(* IEC 61131-3 sources: plc-st-coding-agent/progress/f14_agent_v2/release/datasets/public/tests, 20 files *)

(* ---- public-easy-01.reference.st ---- *)
(* 参考解：Automated filling line control（清洗 -> 灌装 -> 压盖 -> 包装 -> 完成灯 -> 取瓶复位）
   工序号用内部状态 stepNo 表示：0=空闲 1=清洗 2=灌装 3=压盖 4=包装 5=完成。
   只用接口变量做输出，“工序启动后保持运行”由 stepNo 只增不减保证。 *)
FUNCTION_BLOCK FB_FillingLine
VAR_INPUT
    bottleSensor : BOOL;            (* 瓶子到位检测 *)
    cleaningConfirmButton : BOOL;   (* 清洗完成确认 *)
    fillingConfirmButton : BOOL;    (* 灌装完成确认 *)
    cappingConfirmButton : BOOL;    (* 压盖完成确认 *)
    packingConfirmButton : BOOL;    (* 包装完成确认 *)
    finishedButton : BOOL;          (* 取走瓶子确认 *)
END_VAR
VAR_OUTPUT
    Pump_Motor : BOOL;              (* 清洗泵 *)
    Filling_Valve : BOOL;           (* 灌装阀 *)
    Capping_Machine : BOOL;         (* 压盖机 *)
    Packing_Machine : BOOL;         (* 包装机 *)
    Completion_Light : BOOL;        (* 包装完成指示灯 *)
END_VAR
VAR
    stepNo : INT;                   (* 当前工序号，0=空闲 *)
END_VAR

(* R1: 检测到瓶子就启动清洗泵（stepNo 1），此后 stepNo 不回退，泵持续工作 *)
IF bottleSensor AND (stepNo = 0) THEN
    stepNo := 1;
END_IF

(* R2..R5: 每道工序由“上一道工序完成”的确认按钮推进；只接受当拍工序的确认，
   因此误按后道工序的按钮不会跳步，而且机器一旦启动就保持运行 *)
IF (stepNo = 1) AND cleaningConfirmButton THEN
    stepNo := 2;
ELSIF (stepNo = 2) AND fillingConfirmButton THEN
    stepNo := 3;
ELSIF (stepNo = 3) AND cappingConfirmButton THEN
    stepNo := 4;
ELSIF (stepNo = 4) AND packingConfirmButton THEN
    stepNo := 5;
END_IF

(* R6: 取走瓶子 -> 灭灯并整线复位，准备下一循环 *)
IF finishedButton THEN
    stepNo := 0;
END_IF

(* 各执行机构的输出：由工序号唯一决定，故“启动即保持” *)
Pump_Motor := (stepNo >= 1);
Filling_Valve := (stepNo >= 2);
Capping_Machine := (stepNo >= 3);
Packing_Machine := (stepNo >= 4);
Completion_Light := (stepNo = 5);
END_FUNCTION_BLOCK

(* ---- public-easy-02.reference.st ---- *)
(* 参考解：Dual-word edge detection（DWORD 逐位上升沿/下降沿）
   prevValue 保存上一拍的输入值，声明初值为 0（PLC 上电瞬间存储区为 0），
   因此第 1 拍等价于“相对全 0 的边沿检测”，与需求“比较两个连续的 DWORD”一致。 *)
FUNCTION_BLOCK FB_DualWordEdge
VAR_INPUT
    value : DWORD;                  (* 每个周期检查的输入字 *)
END_VAR
VAR_OUTPUT
    hasChanged : BOOL;              (* 有无任何位变化 *)
    hasRisingEdges : BOOL;          (* 有无上升沿 *)
    risingBits : DWORD;             (* 上升沿位流：某位本拍由 0 变 1 则为 1 *)
    noOfRisingBits : USINT;         (* 上升沿位数 *)
    hasFallingEdges : BOOL;         (* 有无下降沿 *)
    fallingBits : DWORD;            (* 下降沿位流：某位本拍由 1 变 0 则为 1 *)
    noOfFallingBits : USINT;        (* 下降沿位数 *)
END_VAR
VAR
    prevValue : DWORD;              (* 上一拍的输入值 *)
    tmpBits : DWORD;                (* 统计位数的移位暂存 *)
    bitCount : USINT;               (* 统计结果暂存 *)
    i : INT;                        (* 循环变量 *)
END_VAR

(* R1/R2: 按位求差。NOT 对整数是 32 位按位取反，与 DWORD 宽度一致。
   IEC 的 AND/OR 两侧都是整数时按位运算，所以这里不会退化成逻辑运算。 *)
risingBits := value AND NOT prevValue;
fallingBits := prevValue AND NOT value;

(* R3: 是否变化，以及两类边沿是否存在 *)
hasChanged := (risingBits <> 0) OR (fallingBits <> 0);
hasRisingEdges := risingBits <> 0;
hasFallingEdges := fallingBits <> 0;

(* R4: 上升沿位数——逐位右移数 1 的个数（32 位，故循环 32 次） *)
bitCount := 0;
tmpBits := risingBits;
FOR i := 1 TO 32 DO
    IF (tmpBits AND 1) <> 0 THEN
        bitCount := bitCount + 1;
    END_IF
    tmpBits := tmpBits SHR 1;
END_FOR
noOfRisingBits := bitCount;

(* R6: 下降沿位数，同一套逐位统计 *)
bitCount := 0;
tmpBits := fallingBits;
FOR i := 1 TO 32 DO
    IF (tmpBits AND 1) <> 0 THEN
        bitCount := bitCount + 1;
    END_IF
    tmpBits := tmpBits SHR 1;
END_FOR
noOfFallingBits := bitCount;

(* R5: 本拍值成为下一拍的“上一拍” *)
prevValue := value;
END_FUNCTION_BLOCK

(* ---- public-easy-03.reference.st ---- *)
(* 参考解：Alarm handling（带回差的高/低限报警 + 参数校验）
   报警输出是锁存量：超过限值才置位，回到“限值 ± 回差”以内才复位（回差防抖）。
   参数非法时置 error 并给出 status，且本次扫描不再评估报警（等价于“退出程序”）。 *)
FUNCTION_BLOCK FB_AlarmHandling
VAR_INPUT
    Value : REAL;                   (* 被监视的输入值 *)
    hiLevel : REAL;                 (* 高限报警值 *)
    loLevel : REAL;                 (* 低限报警值 *)
    hystWindow : REAL;              (* 回差窗口 *)
END_VAR
VAR_OUTPUT
    hiAlarm : BOOL;                 (* 高限报警 *)
    loAlarm : BOOL;                 (* 低限报警 *)
    error : BOOL;                   (* 执行出错 *)
    status : WORD;                  (* 状态码：16#8001 / 16#8002 *)
END_VAR

(* R5: 上下限设置反了（loLevel >= hiLevel）-> error，status=16#8001，退出 *)
IF loLevel >= hiLevel THEN
    error := TRUE;
    status := 16#8001;
(* R6: 回差窗口不比正常范围窄（hystWindow >= hiLevel - loLevel）-> error，status=16#8002 *)
ELSIF hystWindow >= (hiLevel - loLevel) THEN
    error := TRUE;
    status := 16#8002;
ELSE
    error := FALSE;
    status := 16#0000;

    (* R1/R2: 高于高限置位；低于 hiLevel-hystWindow 才复位，中间的过渡带保持原状态 *)
    IF Value > hiLevel THEN
        hiAlarm := TRUE;
    ELSIF Value < (hiLevel - hystWindow) THEN
        hiAlarm := FALSE;
    END_IF

    (* R3/R4: 低于低限置位；高于 loLevel+hystWindow 才复位 *)
    IF Value < loLevel THEN
        loAlarm := TRUE;
    ELSIF Value > (loLevel + hystWindow) THEN
        loAlarm := FALSE;
    END_IF
END_IF
END_FUNCTION_BLOCK

(* ---- public-easy-04.reference.st ---- *)
FUNCTION_BLOCK FB
VAR_INPUT
    VISCOSITY_OK : BOOL;
    PASTE_E_STOP_NC : BOOL;
    DebounceTime : TIME;
    CycleTime : TIME;
END_VAR
VAR_OUTPUT
    VFD_RUN : BOOL;
    PUMP_MAINT_DUE : BOOL;
    PUMP_RUNTIME_ACC : LTIME;
END_VAR
VAR
    viscosityDelay : TON;
END_VAR
viscosityDelay(IN := VISCOSITY_OK AND PASTE_E_STOP_NC, PT := DebounceTime);
VFD_RUN := viscosityDelay.Q;
IF VFD_RUN THEN
    PUMP_RUNTIME_ACC := PUMP_RUNTIME_ACC + TIME_TO_LTIME(CycleTime);
END_IF;
PUMP_MAINT_DUE := PUMP_RUNTIME_ACC >= LTIME#500h;
END_FUNCTION_BLOCK

(* ---- public-easy-05.reference.st ---- *)
FUNCTION_BLOCK FB_WeldGapAlarm
VAR_INPUT
    Gap_Exceeded : BOOL;
    Weld_E_Stop_NC : BOOL;
    DebounceTime : TIME;
END_VAR
VAR_OUTPUT
    Operator_Alert : BOOL;
    Weld_Soft_Start_Active : BOOL;
END_VAR
VAR
    startupDelay : TON;
    gapDelay : TON;
END_VAR
startupDelay(IN := TRUE, PT := T#5s);
Weld_Soft_Start_Active := NOT startupDelay.Q;
gapDelay(IN := startupDelay.Q AND Weld_E_Stop_NC AND Gap_Exceeded, PT := DebounceTime);
Operator_Alert := gapDelay.Q;
END_FUNCTION_BLOCK

(* ---- public-easy-06.reference.st ---- *)
FUNCTION_BLOCK FB_AerationBlower
VAR_INPUT
    DO_LOW : BOOL;
    AERATION_E_STOP_NC : BOOL;
END_VAR
VAR_OUTPUT
    BLOWER_RUN : BOOL;
    AERATION_BLOWER_CYCLE_COUNT : UINT;
END_VAR
VAR
    startDelay : TON;
    wasRunning : BOOL;
END_VAR
startDelay(IN := DO_LOW AND AERATION_E_STOP_NC, PT := T#5s);
BLOWER_RUN := startDelay.Q;
IF BLOWER_RUN AND NOT wasRunning AND AERATION_BLOWER_CYCLE_COUNT < 65535 THEN
    AERATION_BLOWER_CYCLE_COUNT := AERATION_BLOWER_CYCLE_COUNT + 1;
END_IF;
wasRunning := BLOWER_RUN;
END_FUNCTION_BLOCK

(* ---- public-hard-01.reference.st ---- *)
(*
    public-hard-01  Material Proportioning Process Control
    参考解：单个 FUNCTION_BLOCK。接口名与数据类型严格照抄 variables。

    平台说明（公共题制作约定 §7）：
      * 无 TON / R_TRIG，按钮的上升沿用显式边沿
            e := btn AND NOT prev;  prev := btn;
        在扫描末尾统一滚动 prev，避免同拍重复触发。
      * "液位达到 N cm" 用 levelSensor >= N 判断（液位单调上升的语义）。
      * 时间类原语里没有可用的定时器，本题流程全部由 levelSensor / 完成信号推进。

    本文件用 (* R1: ... *) 形式标注需求编号，逐条对应 requirements。
*)
FUNCTION_BLOCK FB_MaterialProportioning
VAR_INPUT
    estop : BOOL;             (* R1 急停：FALSE = 触发 *)
    opeMode : BOOL;           (* R2/R4 运行方式：FALSE = 手动，TRUE = 自动 *)
    valveAStart : BOOL;       (* 手动按钮（上升沿启停） *)
    valveBStart : BOOL;
    valveCStart : BOOL;
    valveDStart : BOOL;
    mixMotorStart : BOOL;
    autoStart : BOOL;         (* 自动流程启动按钮（上升沿） *)
    processMode : BOOL;       (* R5 FALSE = 直接混合；TRUE = 先进 C 到 100cm 再混合 *)
    levelSensor : INT;        (* 液位传感器，单位 cm *)
    mixMotorComplete : BOOL;  (* R6 混合完成信号 *)
END_VAR
VAR_OUTPUT
    valveARun : BOOL;
    valveBRun : BOOL;
    valveCRun : BOOL;
    valveDRun : BOOL;
    mixMotorRun : BOOL;
END_VAR
VAR
    (* 自动流程步序：0 空闲 / 10 进料 A / 20 进料 B / 35 进料 C / 40 混合 / 50 完成 *)
    state : INT;
    (* 各按钮与运行方式上一拍的值（显式边沿用） *)
    prevAutoStart : BOOL;
    prevValveAStart : BOOL;
    prevValveBStart : BOOL;
    prevValveCStart : BOOL;
    prevValveDStart : BOOL;
    prevMixMotorStart : BOOL;
    prevOpeMode : BOOL;
    (* 手动模式下五个设备的启停记忆 *)
    manA : BOOL;
    manB : BOOL;
    manC : BOOL;
    manD : BOOL;
    manMix : BOOL;
END_VAR

(* R1: 急停最高优先级——estop=FALSE 时所有设备立即停机，
   并复位自动流程与手动记忆；急停解除后不会自动续跑，必须重新启动。 *)
IF NOT estop THEN
    state := 0;
    manA := FALSE;
    manB := FALSE;
    manC := FALSE;
    manD := FALSE;
    manMix := FALSE;
    valveARun := FALSE;
    valveBRun := FALSE;
    valveCRun := FALSE;
    valveDRun := FALSE;
    mixMotorRun := FALSE;

(* R2: 手动模式——五个设备各自由对应按钮的上升沿翻转（启/停）。
   R3: 只认上升沿：按住不放不会反复翻转；释放后保持当前状态。 *)
ELSIF NOT opeMode THEN
    (* 从自动切到手动的那一拍：放弃自动流程，手动记忆全部复位（需求未规定，
       取最安全侧，见文件末尾"需求未覆盖处"说明）。 *)
    IF prevOpeMode THEN
        state := 0;
        manA := FALSE;
        manB := FALSE;
        manC := FALSE;
        manD := FALSE;
        manMix := FALSE;
    END_IF
    IF valveAStart AND NOT prevValveAStart THEN
        manA := NOT manA;
    END_IF
    IF valveBStart AND NOT prevValveBStart THEN
        manB := NOT manB;
    END_IF
    IF valveCStart AND NOT prevValveCStart THEN
        manC := NOT manC;
    END_IF
    IF valveDStart AND NOT prevValveDStart THEN
        manD := NOT manD;
    END_IF
    IF mixMotorStart AND NOT prevMixMotorStart THEN
        manMix := NOT manMix;
    END_IF
    valveARun := manA;
    valveBRun := manB;
    valveCRun := manC;
    valveDRun := manD;
    mixMotorRun := manMix;

(* R4/R5/R6: 自动模式——按工艺步序推进设备，手动按钮被忽略。 *)
ELSE
    (* 刚进入自动模式：自动流程从头开始，手动残留输出全部关断。 *)
    IF NOT prevOpeMode THEN
        state := 0;
        valveARun := FALSE;
        valveBRun := FALSE;
        valveCRun := FALSE;
        valveDRun := FALSE;
        mixMotorRun := FALSE;
    END_IF

    CASE state OF
        0:  (* 空闲：等待 autoStart 上升沿 *)
            valveARun := FALSE;
            valveBRun := FALSE;
            valveCRun := FALSE;
            valveDRun := FALSE;
            mixMotorRun := FALSE;
            (* R4: 按 autoStart 启动自动流程，先开阀 A *)
            IF autoStart AND NOT prevAutoStart THEN
                state := 10;
                valveARun := TRUE;
            END_IF

        10: (* 进料 A：液位到 50cm 关 A、开 B *)
            valveARun := TRUE;
            valveBRun := FALSE;
            valveCRun := FALSE;
            valveDRun := FALSE;
            mixMotorRun := FALSE;
            IF levelSensor >= 50 THEN
                valveARun := FALSE;
                valveBRun := TRUE;
                state := 20;
            END_IF

        20: (* 进料 B：液位到 80cm 关 B；随后按 processMode 决定下一步 *)
            valveARun := FALSE;
            valveBRun := TRUE;
            valveCRun := FALSE;
            valveDRun := FALSE;
            mixMotorRun := FALSE;
            IF levelSensor >= 80 THEN
                valveBRun := FALSE;
                IF processMode THEN
                    (* R5(true): 先开 C 继续进料到 100cm *)
                    valveCRun := TRUE;
                    state := 35;
                ELSE
                    (* R5(false): 不进 C，直接启动混合电机 *)
                    mixMotorRun := TRUE;
                    state := 40;
                END_IF
            END_IF

        35: (* 进料 C：液位到 100cm 关 C、启动混合电机 *)
            valveARun := FALSE;
            valveBRun := FALSE;
            valveCRun := TRUE;
            valveDRun := FALSE;
            mixMotorRun := FALSE;
            IF levelSensor >= 100 THEN
                valveCRun := FALSE;
                mixMotorRun := TRUE;
                state := 40;
            END_IF

        40: (* 混合中：收到混合完成信号 → 停电机、开 D、流程结束 *)
            valveARun := FALSE;
            valveBRun := FALSE;
            valveCRun := FALSE;
            valveDRun := FALSE;
            mixMotorRun := TRUE;
            IF mixMotorComplete THEN
                mixMotorRun := FALSE;
                valveDRun := TRUE;
                state := 50;
            END_IF

        50: (* 完成：D 保持开启把料送出；再次 autoStart 开始新一周期 *)
            valveARun := FALSE;
            valveBRun := FALSE;
            valveCRun := FALSE;
            valveDRun := TRUE;
            mixMotorRun := FALSE;
            IF autoStart AND NOT prevAutoStart THEN
                valveDRun := FALSE;
                valveARun := TRUE;
                state := 10;
            END_IF
    END_CASE
END_IF

(* 边沿记忆统一在扫描末尾滚动（顺序不可提前，见约定 §7）。 *)
prevAutoStart := autoStart;
prevValveAStart := valveAStart;
prevValveBStart := valveBStart;
prevValveCStart := valveCStart;
prevValveDStart := valveDStart;
prevMixMotorStart := mixMotorStart;
prevOpeMode := opeMode;

(*
  需求未覆盖处的取舍（均为最安全侧，且已由 test_cases 覆盖其行为）：
  1) 运行方式切换：自动→手动或手动→自动时，当前流程被中止、输出全部关断，
     不会在切换后残留上一模式的设备动作；自动模式要从步序 0 重新 autoStart。
  2) 自动流程进行中再次按 autoStart 被忽略（按键只对步序 0 / 50 有效），
     避免运行中反复重启流程。
  3) 自动完成后阀 D 保持开启（"open valve D, and the automatic process ends"），
     直到下一次 autoStart 开始新周期或急停触发。
  4) 步序 0 与各步都显式给全部输出赋值，保证同一扫描周期内输出不残留上一步的值。
*)
END_FUNCTION_BLOCK

(* ---- public-hard-02.reference.st ---- *)
(* public-hard-02 Flexible Processing Control
   1# 上料 / 2#~4# 加工 / 5# 出库。工序序列由 processSequence + processLength 给出，
   processLength 从 processSequence[1] 起算，末项由 caller 保证是 5# 出库站。
   内部状态机 phase：0=空闲/待料，1=输送中，2=等当前加工工位完成信号。 *)

FUNCTION_BLOCK FB
VAR_INPUT
    processLength : USINT;
    sensor1 : BOOL;
    sensor2 : BOOL;
    sensor3 : BOOL;
    sensor4 : BOOL;
    sensor5 : BOOL;
    station1Start : BOOL;
    station2Complete : BOOL;
    station3Complete : BOOL;
    station4Complete : BOOL;
    processSequence : ARRAY[1..8] OF USINT;
END_VAR
VAR_OUTPUT
    conveyorLeft : BOOL;
    conveyorRight : BOOL;
END_VAR
VAR
    phase : INT;          (* 0 空闲；1 输送中；2 等加工完成 *)
    idx : INT;            (* 当前执行到 processSequence 的第几项 *)
    curStation : INT;     (* 产品当前所在工位 *)
    dstStation : INT;     (* 本段输送的目标工位 *)
    lenNow : INT;
    dstOK : BOOL;
    arrived : BOOL;
    startEdge : BOOL;
    startPrev : BOOL;
    compEdge : BOOL;
    comp2Prev : BOOL;
    comp3Prev : BOOL;
    comp4Prev : BOOL;
END_VAR

(* R1/R2: 启动按钮上升沿 + 1# 有料才启动；序列长度必须落在 1..8 *)
startEdge := station1Start AND NOT startPrev;
startPrev := station1Start;
lenNow := processLength;

(* 加工完成信号按上升沿消费；每拍都刷新历史值，避免边沿被相位切换吃掉 *)
compEdge := FALSE;
IF phase = 2 THEN
    IF curStation = 2 THEN
        compEdge := station2Complete AND NOT comp2Prev;
    ELSIF curStation = 3 THEN
        compEdge := station3Complete AND NOT comp3Prev;
    ELSIF curStation = 4 THEN
        compEdge := station4Complete AND NOT comp4Prev;
    END_IF;
END_IF;
comp2Prev := station2Complete;
comp3Prev := station3Complete;
comp4Prev := station4Complete;

conveyorLeft := FALSE;
conveyorRight := FALSE;

(* R1: 上料工位有料 + 按下启动 → 查第一个工序号，当拍就启动输送带 *)
IF phase = 0 THEN
    IF sensor1 AND startEdge THEN
        IF (lenNow >= 1) AND (lenNow <= 8) THEN
            dstStation := processSequence[1];
            dstOK := (dstStation >= 2) AND (dstStation <= 5);
            IF dstOK THEN
                idx := 1;
                curStation := 1;
                phase := 1;
            END_IF;
        END_IF;
    END_IF;
END_IF;

(* R4: 收到当前工位完成信号 → 查下一个工序号，当拍转向继续输送 *)
IF phase = 2 THEN
    IF compEdge THEN
        idx := idx + 1;
        IF (idx > lenNow) OR (idx > 8) THEN
            (* 非法序列（末项不是 5#）的保护：不再读数组下标，直接停机 *)
            phase := 0;
        ELSE
            dstStation := processSequence[idx];
            dstOK := (dstStation >= 2) AND (dstStation <= 5);
            IF dstOK THEN
                phase := 1;
            ELSE
                phase := 0;
            END_IF;
        END_IF;
    END_IF;
END_IF;

(* R3/R5: 按 "目标工位 vs 当前工位" 决定方向；只看目标工位传感器判到位 *)
IF phase = 1 THEN
    IF dstStation > curStation THEN
        conveyorRight := TRUE;
    ELSIF dstStation < curStation THEN
        conveyorLeft := TRUE;
    END_IF;
    arrived := FALSE;
    IF dstStation = 2 THEN
        arrived := sensor2;
    ELSIF dstStation = 3 THEN
        arrived := sensor3;
    ELSIF dstStation = 4 THEN
        arrived := sensor4;
    ELSIF dstStation = 5 THEN
        arrived := sensor5;
    END_IF;
    IF arrived THEN
        conveyorLeft := FALSE;
        conveyorRight := FALSE;
        curStation := dstStation;
        IF dstStation = 5 THEN
            (* R5: 送到 5# 出库站，一个产品的流程结束 *)
            phase := 0;
        ELSE
            (* R4: 停在该工位，等它给出加工完成信号 *)
            phase := 2;
        END_IF;
    END_IF;
END_IF;
END_FUNCTION_BLOCK

(* ---- public-hard-03.reference.st ---- *)
(*
  Recipe Management System — 参考解（public-hard-03）

  配方库 recipe 是 VAR_IN_OUT 的结构体数组，最多 10 条，recipeID = 0 表示空槽；
  四个请求信号取上升沿，因此一个请求只执行一次（电平保持不会重复执行）。

  需求编号（对应 requirements 的 Notes）：
    R2  查询：号码不存在 -> error=TRUE & status=16#8001；存在 -> 输出到 recipeQueryResult
    R3  新增：号码重复 -> 16#8002；无空槽 -> 16#8003；否则存到下标最小的空槽
    R4  删除：号码不存在 -> 16#8004；存在 -> 把该槽的 recipeID 置 0
    R5  修改：号码不存在 -> 16#8005；存在 -> 用 recipeIn 覆盖该槽
  另有 R1：配方字段 recipeID/ingredientType/ingredientRatio/productionTemperature。

  两处按需求原文做的判定口径（都写在下面的注释里）：
    * 0 号不是合法配方号：查询/删除/修改 0 号一律按"号码不存在"处理；
    * 新增时号码与本库任何一条 recipeID 相同即算重复，因此 0 号会与空槽的 0 相撞，
      在还有空槽时报 16#8002（R3 的判定顺序本来就是"先查重复、再查空槽"）。
*)

TYPE ST_Recipe :
STRUCT
  recipeID : INT;                (* 配方号，0 = 空槽 *)
  ingredientType : INT;          (* 原料类型 *)
  ingredientRatio : REAL;        (* 原料配比 *)
  productionTemperature : REAL;  (* 生产温度 *)
END_STRUCT
END_TYPE

FUNCTION_BLOCK FB
VAR_INPUT
  addRecipe : BOOL;              (* R3 新增请求 *)
  deleteRecipe : BOOL;           (* R4 删除请求 *)
  modifyRecipe : BOOL;           (* R5 修改请求 *)
  queryRecipe : BOOL;            (* R2 查询请求 *)
  recipeIn : ST_Recipe;          (* 请求携带的配方 *)
END_VAR
VAR_OUTPUT
  recipeAdded : BOOL;            (* 新增成功指示，只在执行成功那一拍为 TRUE *)
  recipeDeleted : BOOL;          (* 删除成功指示 *)
  recipeModified : BOOL;         (* 修改成功指示 *)
  recipeQueryResult : ST_Recipe; (* 查询结果，只在查询成功时更新 *)
  error : BOOL;                  (* 出错指示 *)
  status : WORD;                 (* 状态码，0 = 正常 *)
END_VAR
VAR_IN_OUT
  recipe : ARRAY[1..10] OF ST_Recipe;   (* 配方库 *)
END_VAR
VAR
  i : INT;
  hitIdx : INT;                  (* 命中槽，0 = 没命中 *)
  freeIdx : INT;                 (* 下标最小的空槽，0 = 库已满 *)
  dup : BOOL;                    (* 新增时号码重复 *)
  qEdge : BOOL;  qPrev : BOOL;   (* R2 请求上升沿 *)
  aEdge : BOOL;  aPrev : BOOL;   (* R3 *)
  dEdge : BOOL;  dPrev : BOOL;   (* R4 *)
  mEdge : BOOL;  mPrev : BOOL;   (* R5 *)
END_VAR

(* 成功指示与状态码都是"拍"语义：每个周期先清零，只在执行请求的那一拍置位 *)
recipeAdded := FALSE;
recipeDeleted := FALSE;
recipeModified := FALSE;
error := FALSE;
status := 16#0000;

(* 请求信号取上升沿：按钮保持为 TRUE 时不会每个扫描周期都重做一遍 *)
qEdge := queryRecipe AND NOT qPrev;
qPrev := queryRecipe;
aEdge := addRecipe AND NOT aPrev;
aPrev := addRecipe;
dEdge := deleteRecipe AND NOT dPrev;
dPrev := deleteRecipe;
mEdge := modifyRecipe AND NOT mPrev;
mPrev := modifyRecipe;

(* 在库里找 recipeIn 的配方号；0 号是"空槽标记"而不是配方，一律当不存在 *)
hitIdx := 0;
IF recipeIn.recipeID <> 0 THEN
  FOR i := 1 TO 10 DO
    IF (hitIdx = 0) AND (recipe[i].recipeID = recipeIn.recipeID) THEN
      hitIdx := i;
    END_IF
  END_FOR
END_IF

(* 下标最小的空槽，供 R3 的落地位置使用 *)
freeIdx := 0;
FOR i := 1 TO 10 DO
  IF (freeIdx = 0) AND (recipe[i].recipeID = 0) THEN
    freeIdx := i;
  END_IF
END_FOR

(* 四条需求是各自并列的规则：每个请求在自己的上升沿被执行一次，互不吞并 *)
IF qEdge THEN
  (* R2 查询 *)
  IF hitIdx = 0 THEN
    error := TRUE;
    status := 16#8001;
  ELSE
    recipeQueryResult.recipeID := recipe[hitIdx].recipeID;
    recipeQueryResult.ingredientType := recipe[hitIdx].ingredientType;
    recipeQueryResult.ingredientRatio := recipe[hitIdx].ingredientRatio;
    recipeQueryResult.productionTemperature := recipe[hitIdx].productionTemperature;
  END_IF
END_IF

IF aEdge THEN
  (* R3 新增：先查重号，再查空槽 *)
  dup := FALSE;
  FOR i := 1 TO 10 DO
    IF (NOT dup) AND (recipe[i].recipeID = recipeIn.recipeID) THEN
      dup := TRUE;
    END_IF
  END_FOR
  IF dup THEN
    error := TRUE;
    status := 16#8002;
  ELSIF freeIdx = 0 THEN
    error := TRUE;
    status := 16#8003;
  ELSE
    recipe[freeIdx].recipeID := recipeIn.recipeID;
    recipe[freeIdx].ingredientType := recipeIn.ingredientType;
    recipe[freeIdx].ingredientRatio := recipeIn.ingredientRatio;
    recipe[freeIdx].productionTemperature := recipeIn.productionTemperature;
    recipeAdded := TRUE;
  END_IF
END_IF

IF dEdge THEN
  (* R4 删除：只清配方号，槽位立即可以被后续新增复用 *)
  IF hitIdx = 0 THEN
    error := TRUE;
    status := 16#8004;
  ELSE
    recipe[hitIdx].recipeID := 0;
    recipeDeleted := TRUE;
  END_IF
END_IF

IF mEdge THEN
  (* R5 修改：整条配方用 recipeIn 覆盖（结构体不能整体赋值，只能逐字段） *)
  IF hitIdx = 0 THEN
    error := TRUE;
    status := 16#8005;
  ELSE
    recipe[hitIdx].recipeID := recipeIn.recipeID;
    recipe[hitIdx].ingredientType := recipeIn.ingredientType;
    recipe[hitIdx].ingredientRatio := recipeIn.ingredientRatio;
    recipe[hitIdx].productionTemperature := recipeIn.productionTemperature;
    recipeModified := TRUE;
  END_IF
END_IF

END_FUNCTION_BLOCK

(* ---- public-hard-04.reference.st ---- *)
(*
  FIFO Circular Queue with VARIANT Storage — 参考解（public-hard-04）

  容量与元素类型都来自调用方数组 buffer（VARIANT 里的真实数组，容量 = 数组长度），
  内部只维护 head（队头下标，1 起）与 count（有效元素个数）；tail 由二者算出，
  head/tail/count 都不出现在接口上（R6）。

  需求编号：
    R1  入队请求上升沿 -> 队列未满时把当前 item 追加到队尾
    R2  出队请求上升沿 -> 队列非空时移除队首并把该值写回 item
    R3  reset=TRUE 清空队列、elementCount=0，且优先于入队/出队
    R4  elementCount 输出当前有效元素个数（0 空、等于容量为满）
    R5  空队出队/满队入队要拒绝：队列与 item 保持不变，status 说明原因
    R6  首次调用时队列为空；head/tail 等内部状态不出现在接口上
*)

FUNCTION_BLOCK FB
VAR_INPUT
  enqueue : BOOL;                (* R1 入队请求，一个上升沿执行一次 *)
  dequeue : BOOL;                (* R2 出队请求，一个上升沿执行一次 *)
  reset : BOOL;                  (* R3 复位，优先于入队/出队 *)
END_VAR
VAR_OUTPUT
  elementCount : DINT;           (* R4 当前有效元素个数 *)
  status : WORD;                 (* R5 16#0000 / 16#8001 / 16#8002 *)
END_VAR
VAR_IN_OUT
  item : VARIANT;                (* 入队时读取；出队成功时写回被移除的队首值 *)
  buffer : VARIANT;              (* 队列存储，容量 = 数组实际长度 *)
END_VAR
VAR
  cap : DINT;                    (* 本拍看到的容量 *)
  count : DINT;                  (* 有效元素个数，不放接口（R6） *)
  head : DINT;                   (* 队头下标（1 起） *)
  tail : DINT;                   (* 队尾插入位置（由 head+count 算出） *)
  enEdge : BOOL;  enPrev : BOOL; (* R1 上升沿 *)
  deEdge : BOOL;  dePrev : BOOL; (* R2 上升沿 *)
END_VAR

(* 容量每拍从调用方数组重新取：数组换长度时行为随之改变 *)
cap := UPPER_BOUND(buffer, 1) - LOWER_BOUND(buffer, 1) + 1;

(* 内部下标兜底：首次调用 / 复位后 head 一定落在 1..cap *)
IF count < 0 THEN
  count := 0;
END_IF
IF head < 1 THEN
  head := 1;
END_IF

(* 上升沿：一次请求只执行一次，按住不放不会重复入队/出队 *)
enEdge := enqueue AND NOT enPrev;
enPrev := enqueue;
deEdge := dequeue AND NOT dePrev;
dePrev := dequeue;

(* 状态码是"拍"语义：每拍先回到 16#0000，只有被拒绝的那一拍才置错误码 *)
status := 16#0000;

IF reset THEN
  (* R3 复位优先：同时到来的入队/出队请求被丢弃，只清空队列 *)
  count := 0;
  head := 1;
ELSIF enEdge THEN
  (* R1 入队 *)
  IF (cap <= 0) OR (count >= cap) THEN
    status := 16#8002;         (* R5 满队（容量为 0 的数组也按"装不下"拒绝） *)
  ELSE
    IF count > cap - head THEN
      tail := count - (cap - head);
    ELSE
      tail := head + count;    (* 此分支已知和不超过 cap，适用于 DINT 极值容量 *)
    END_IF
    buffer[LOWER_BOUND(buffer, 1) + (tail - 1)] := item;      (* VARIANT 元素写入：类型由数组元素决定 *)
    count := count + 1;
  END_IF
ELSIF deEdge THEN
  (* R2 出队 *)
  IF count <= 0 THEN
    status := 16#8001;         (* R5 空队，item 保持原值 *)
  ELSE
    item := buffer[LOWER_BOUND(buffer, 1) + (head - 1)];      (* 被移除的队首值写回 item *)
    IF head = cap THEN
      head := 1;
    ELSE
      head := head + 1;
    END_IF
    count := count - 1;
  END_IF
END_IF

(* R4 *)
elementCount := count;

END_FUNCTION_BLOCK

(* ---- public-hard-05.reference.st ---- *)
(*
  Mechanical Arm Control — 参考解（public-hard-05）

  六动作：下/上/左/右/抓/放；四模式：手动/单步/单循环/连续（调用方保证互斥）。
  EmergencyStop 为反逻辑：FALSE = 急停触发，TRUE = 无急停。

  需求编号：
    R1  手动模式：按住按钮且未到位才动作，到位即停，松手即停
    R2  单步模式：按一次 Start 执行预置程序的"下一个"动作，动作完成即停等下一次确认
        预置程序：①下 ②抓 ③上 ④右 ⑤下 ⑥放 ⑦上 ⑧左，第 8 步之后回到第 1 步
    R3  单循环模式：按 Start 自动完成一整套搬运循环，最后一动（回左）到位后停在左上
    R4  连续模式：按 Start 后反复执行 R3 的搬运循环，不停
    R5  急停：任何模式任何时刻都能立刻停掉所有动作（FALSE 有效）；解除后从冻结的位置继续
        模式切换也立刻停掉自动动作，程序步回到起点
    R6  抓/放的完成反馈分别是 GripLimitSwitch / ReleaseLimitSwitch
*)

FUNCTION_BLOCK FB
VAR_INPUT
  (* 四模式，调用方保证同一时刻只有一个为 TRUE（本实现对同时为 TRUE 的容错 = 取高者） *)
  ManualMode : BOOL;             (* R1 *)
  SingleStepMode : BOOL;         (* R2 *)
  SingleCycleMode : BOOL;        (* R3 *)
  ContinuousMode : BOOL;         (* R4 *)
  EmergencyStop : BOOL;          (* R5 FALSE = 急停 *)
  Start : BOOL;                  (* R2/R3/R4 每按一次算一条指令 *)
  DownButton : BOOL;             (* R1 *)
  UpButton : BOOL;               (* R1 *)
  LeftButton : BOOL;             (* R1 *)
  RightButton : BOOL;            (* R1 *)
  GripButton : BOOL;             (* R1 *)
  ReleaseButton : BOOL;          (* R1 *)
  DownLimitSwitch : BOOL;        (* 到位反馈 *)
  UpLimitSwitch : BOOL;
  LeftLimitSwitch : BOOL;
  RightLimitSwitch : BOOL;
  GripLimitSwitch : BOOL;        (* R6 抓完成 *)
  ReleaseLimitSwitch : BOOL;     (* R6 放完成 *)
END_VAR
VAR_OUTPUT
  MoveDown : BOOL;
  MoveUp : BOOL;
  MoveLeft : BOOL;
  MoveRight : BOOL;
  ActivateGrip : BOOL;
  ActivateRelease : BOOL;
END_VAR
VAR
  startEdge : BOOL;              (* Start 上升沿 *)
  startPrev : BOOL;
  modeNow : INT;                 (* 本拍模式号 0 无 / 1 手动 / 2 单步 / 3 单循环 / 4 连续 *)
  modePrev : INT;
  fsStep : INT;                  (* 预置程序的当前步 1..8；0 = 未开始或本轮已结束 *)
  fsActive : BOOL;               (* 自动程序是否正在执行某个动作 *)
  fsDone : BOOL;                 (* 当前步的到位条件是否已满足 *)
  guard : INT;                   (* 每拍最多推进 8 步，防止一拍扫完多圈 *)
END_VAR

(* 每拍先把六个动作输出清零，后面按模式/状态逐位置位：急停或无模式时自然全 0（R5） *)
MoveDown := FALSE;
MoveUp := FALSE;
MoveLeft := FALSE;
MoveRight := FALSE;
ActivateGrip := FALSE;
ActivateRelease := FALSE;

(* 上升沿：按一次 Start 只发一条指令，按住不放不会连发 *)
startEdge := Start AND NOT startPrev;
startPrev := Start;

(* 模式号：四模式互斥由调用方保证；若同时为 TRUE 按 手动 > 单步 > 单循环 > 连续 取高者 *)
modeNow := 0;
IF ContinuousMode THEN
  modeNow := 4;
END_IF
IF SingleCycleMode THEN
  modeNow := 3;
END_IF
IF SingleStepMode THEN
  modeNow := 2;
END_IF
IF ManualMode THEN
  modeNow := 1;
END_IF

(* R5 模式切换：立刻停掉自动动作并把程序步清回起点，等新模式的指令 *)
IF modeNow <> modePrev THEN
  fsActive := FALSE;
  fsStep := 0;
  fsDone := FALSE;
END_IF
modePrev := modeNow;

IF NOT EmergencyStop THEN
  (* R5 急停压过一切：六个动作全部保持 0，程序步冻结（解除急停后从冻结点继续） *)
  fsDone := FALSE;
ELSIF modeNow = 1 THEN
  (* R1 手动模式：按住按钮且未到位才动作；一对互补按钮同按视为无效（不许同时动作） *)
  IF DownButton AND (NOT DownLimitSwitch) AND (NOT UpButton) THEN
    MoveDown := TRUE;
  END_IF
  IF UpButton AND (NOT UpLimitSwitch) AND (NOT DownButton) THEN
    MoveUp := TRUE;
  END_IF
  IF LeftButton AND (NOT LeftLimitSwitch) AND (NOT RightButton) THEN
    MoveLeft := TRUE;
  END_IF
  IF RightButton AND (NOT RightLimitSwitch) AND (NOT LeftButton) THEN
    MoveRight := TRUE;
  END_IF
  IF GripButton AND (NOT GripLimitSwitch) AND (NOT ReleaseButton) THEN
    ActivateGrip := TRUE;
  END_IF
  IF ReleaseButton AND (NOT ReleaseLimitSwitch) AND (NOT GripButton) THEN
    ActivateRelease := TRUE;
  END_IF
ELSIF (modeNow = 2) OR (modeNow = 3) OR (modeNow = 4) THEN
  (* R2/R3/R4 自动程序 *)
  IF startEdge AND (NOT fsActive) THEN
    IF modeNow = 2 THEN
      (* 单步：接着上次停下的位置继续；还没开始过就从第 1 步起 *)
      IF fsStep < 1 THEN
        fsStep := 1;
      END_IF
    ELSE
      (* 单循环 / 连续：每次启动都从第 1 步（下）重新开始一整轮 *)
      fsStep := 1;
    END_IF
    fsActive := TRUE;
  END_IF

  guard := 0;
  WHILE fsActive AND (guard < 8) DO
    guard := guard + 1;
    fsDone := FALSE;
    (* 预置程序：①下 ②抓 ③上 ④右 ⑤下 ⑥放 ⑦上 ⑧左 *)
    IF fsStep = 1 THEN
      IF DownLimitSwitch THEN fsDone := TRUE; ELSE MoveDown := TRUE; END_IF
    ELSIF fsStep = 2 THEN
      IF GripLimitSwitch THEN fsDone := TRUE; ELSE ActivateGrip := TRUE; END_IF
    ELSIF fsStep = 3 THEN
      IF UpLimitSwitch THEN fsDone := TRUE; ELSE MoveUp := TRUE; END_IF
    ELSIF fsStep = 4 THEN
      IF RightLimitSwitch THEN fsDone := TRUE; ELSE MoveRight := TRUE; END_IF
    ELSIF fsStep = 5 THEN
      IF DownLimitSwitch THEN fsDone := TRUE; ELSE MoveDown := TRUE; END_IF
    ELSIF fsStep = 6 THEN
      IF ReleaseLimitSwitch THEN fsDone := TRUE; ELSE ActivateRelease := TRUE; END_IF
    ELSIF fsStep = 7 THEN
      IF UpLimitSwitch THEN fsDone := TRUE; ELSE MoveUp := TRUE; END_IF
    ELSE
      IF LeftLimitSwitch THEN fsDone := TRUE; ELSE MoveLeft := TRUE; END_IF
    END_IF

    IF NOT fsDone THEN
      (* 本拍动作还没走完：停在当前步，本拍只输出这一个动作 *)
      guard := 8;
    ELSIF modeNow = 4 THEN
      (* R4 连续：本步一完成当拍就进入下一步，第 8 步之后回到第 1 步 *)
      fsStep := fsStep + 1;
      IF fsStep > 8 THEN
        fsStep := 1;
      END_IF
    ELSIF modeNow = 3 THEN
      (* R3 单循环：第 8 步（回左）完成即整轮结束，停在左上等下一次启动 *)
      IF fsStep >= 8 THEN
        fsActive := FALSE;
        fsStep := 0;
      ELSE
        fsStep := fsStep + 1;
      END_IF
    ELSE
      (* R2 单步：一个动作做完就停，等下一次 Start 确认 *)
      fsActive := FALSE;
      fsStep := fsStep + 1;
      IF fsStep > 8 THEN
        fsStep := 1;
      END_IF
    END_IF
  END_WHILE
END_IF

END_FUNCTION_BLOCK

(* ---- public-hard-06.reference.st ---- *)
(*
  Production Control — 参考解（public-hard-06）

  五个工位：上料(Feed) → 清洗(Wash) → 称重(Weight) → 烧结(Firing) → 成品(Output)，
  一台电机负责在工位间传送产品；每个工位一个到位传感器。

  需求编号：
    R1  Mode 开关：FALSE = 手动，TRUE = 自动
    R2  手动模式：ForwardButton 控制正转、ReverseButton 控制反转；正反转必须互锁，不能同时动作
    R3  自动模式：
        a) SensorFeed 检测到料 → 正转送到清洗站 → SensorWash 到位即停 → washComplete 后正转送称重
        b) SensorWeight 到位即停 → weightComplete 后按重量判定：100 ≤ weight ≤ 200 合格
        c) 不合格 → 发出 kick 剔除指令（一拍脉冲），产品被踢出，产线回到等待上料
        d) 合格 → 烧结温度按重量线性映射 100→500、200→550，输出 firingTemp，同时正转送烧结站
        e) SensorFiring 到位即停 → firingComplete 后正转送成品站
        f) SensorOutput 到位即停、CompletionLight 亮；产品被取走（SensorOutput=FALSE）灯灭，回到等待上料
    R4  模式切换：切到手动时自动流程复位（手动接管产线）；切回自动从等待上料重新开始
*)

FUNCTION_BLOCK FB
VAR_INPUT
  Mode : BOOL;                   (* R1 FALSE = 手动，TRUE = 自动 *)
  ForwardButton : BOOL;          (* R2 *)
  ReverseButton : BOOL;          (* R2 *)
  SensorFeed : BOOL;             (* 上料站到位传感器 *)
  SensorWash : BOOL;             (* 清洗站到位传感器 *)
  SensorWeight : BOOL;           (* 称重站到位传感器 *)
  SensorFiring : BOOL;           (* 烧结站到位传感器 *)
  SensorOutput : BOOL;           (* 成品站到位传感器 *)
  washComplete : BOOL;           (* 清洗完成信号 *)
  weightComplete : BOOL;         (* 称重完成信号 *)
  weight : REAL;                 (* 重量值（称重完成时有效） *)
  firingComplete : BOOL;         (* 烧结完成信号 *)
END_VAR
VAR_OUTPUT
  MotorForward : BOOL;           (* 电机正转 *)
  MotorReverse : BOOL;           (* 电机反转（仅手动可用） *)
  kick : BOOL;                   (* 不合格剔除指令 *)
  CompletionLight : BOOL;        (* 成品站完成灯 *)
  firingTemp : REAL;             (* 烧结温度设定值 *)
END_VAR
VAR
  state : INT;                   (* 0 等上料 / 1 送清洗 / 2 等清洗 / 3 送称重 / 4 等称重
                                    5 送烧结 / 6 等烧结 / 7 送成品 / 8 成品站 *)
  modePrev : BOOL;
END_VAR

(* 每拍先清零六个输出：手动/自动互斥由此保证，kick 是脉冲 *)
MotorForward := FALSE;
MotorReverse := FALSE;
kick := FALSE;
CompletionLight := FALSE;

(* R4 模式切换那一拍：自动流程复位，切回自动从"等待上料"重新开始 *)
IF Mode <> modePrev THEN
  state := 0;
END_IF
modePrev := Mode;

IF NOT Mode THEN
  (* R2 手动：两个按钮互锁，同按视为无效（谁都不动） *)
  IF ForwardButton AND (NOT ReverseButton) THEN
    MotorForward := TRUE;
  END_IF
  IF ReverseButton AND (NOT ForwardButton) THEN
    MotorReverse := TRUE;
  END_IF
ELSE
  (* R3 自动流程 *)
  CASE state OF
    0:
      (* 等上料：SensorFeed 检测到料就开始正转送清洗站 *)
      IF SensorFeed THEN
        state := 1;
        MotorForward := TRUE;
      END_IF
    1:
      (* 送到清洗站：到位即停 *)
      IF SensorWash THEN
        state := 2;
      ELSE
        MotorForward := TRUE;
      END_IF
    2:
      (* 等清洗完成 *)
      IF washComplete THEN
        state := 3;
        MotorForward := TRUE;
      END_IF
    3:
      (* 送到称重站：到位即停 *)
      IF SensorWeight THEN
        state := 4;
      ELSE
        MotorForward := TRUE;
      END_IF
    4:
      (* 等称重完成，按 R3b 判定合格与否 *)
      IF weightComplete THEN
        IF (weight >= 100.0) AND (weight <= 200.0) THEN
          (* R3d 合格：100..200 线性映射到 500..550（每 1 个单位重量 0.5 度） *)
          firingTemp := 500.0 + (weight - 100.0) * 0.5;
          state := 5;
          MotorForward := TRUE;
        ELSE
          (* R3c 不合格：剔除，一拍脉冲后回到等待上料；温度保持上一件合格品的值 *)
          kick := TRUE;
          state := 0;
        END_IF
      END_IF
    5:
      (* 送到烧结站：到位即停 *)
      IF SensorFiring THEN
        state := 6;
      ELSE
        MotorForward := TRUE;
      END_IF
    6:
      (* 等烧结完成 *)
      IF firingComplete THEN
        state := 7;
        MotorForward := TRUE;
      END_IF
    7:
      (* 送到成品站：到位即停，完成灯亮 *)
      IF SensorOutput THEN
        state := 8;
        CompletionLight := TRUE;
      ELSE
        MotorForward := TRUE;
      END_IF
    8:
      (* 成品站：产品还在则灯保持亮；被取走则灯灭并回到等待上料 *)
      IF SensorOutput THEN
        CompletionLight := TRUE;
      ELSE
        state := 0;
      END_IF
  ELSE
    state := 0;
  END_CASE
END_IF

END_FUNCTION_BLOCK

(* ---- public-medium-01.reference.st ---- *)
(* 结构体必须显式定义：题目给的是 IN_OUT ARRAY[1..5] OF ST_Pump，
   没有 TYPE 块就读不到字段名，pumpGroup[i].xxx 会被判错。 *)
TYPE ST_Pump :
STRUCT
    priority : INT;    (* 优先级，越大越优先；本 FB 只读 *)
    selection : BOOL;  (* 手动选中状态；本 FB 只读 *)
    RunComd : BOOL;    (* 本 FB 唯一写的字段 *)
END_STRUCT
END_TYPE

FUNCTION_BLOCK FB_MultiPump
VAR_INPUT
    mode : BOOL;   (* FALSE: 手动；TRUE: 自动 *)
    start : BOOL;  (* 启动按钮 *)
    stop : BOOL;   (* 停止按钮：停全部泵 *)
END_VAR
VAR_IN_OUT
    pumpGroup : ARRAY[1..5] OF ST_Pump;
END_VAR
VAR
    i : INT;
    j : INT;
    rank : INT;      (* 第 i 台泵在 5 台里的优先级名次（0 最高） *)
    prioI : INT;
    prioJ : INT;
    inTop3 : BOOL;
END_VAR

(* R4: 停止按钮优先于一切——先无条件把 5 台泵的命令都置 FALSE，
   再进入模式分支；这样 stop 与 start 同时按下时表现为停止。 *)
IF stop THEN
    FOR i := 1 TO 5 DO
        pumpGroup[i].RunComd := FALSE;
    END_FOR

(* R1: 依据 mode 切换运行方式。 *)
ELSIF mode THEN
    (* R3: 自动方式——按 priority 选 3 台（三用两备）。
       不排序、不搬结构体：名次 = 优先级比我高（或同级但下标更小）的台数，
       名次 < 3 即为前三。优先级相同按下标小者优先，保证结果唯一。 *)
    FOR i := 1 TO 5 DO
        rank := 0;
        prioI := pumpGroup[i].priority;
        FOR j := 1 TO 5 DO
            IF j <> i THEN
                prioJ := pumpGroup[j].priority;
                IF (prioJ > prioI) OR ((prioJ = prioI) AND (j < i)) THEN
                    rank := rank + 1;
                END_IF
            END_IF
        END_FOR
        inTop3 := rank < 3;
        (* R2': 自动方式下 start 启动被选中的前 3 台，备用的 2 台必须停机命令 *)
        pumpGroup[i].RunComd := start AND inTop3;
    END_FOR

ELSE
    (* R2: 手动方式——按 selection 逐台控制：选中的泵由 start 启动，
       未选中的泵给停机命令（互斥，不允许两台互相抢）。 *)
    FOR i := 1 TO 5 DO
        pumpGroup[i].RunComd := start AND pumpGroup[i].selection;
    END_FOR
END_IF

END_FUNCTION_BLOCK

(* ---- public-medium-02.reference.st ---- *)
TYPE ST_AnalogChannel :
STRUCT
    enable : BOOL;
    hiLIM : REAL;
    loLIM : REAL;
    bipolar : BOOL;
    measuringMode : INT;
    retVal : WORD;
    outputValue : REAL;
END_STRUCT
END_TYPE

FUNCTION_BLOCK FB
VAR_INPUT
    count : DINT;
END_VAR
VAR_IN_OUT
    analogValues : ARRAY[*] OF INT;
    channels : ARRAY[*] OF ST_AnalogChannel;
END_VAR
VAR
    i : DINT;
    rawBase : DINT;
    channelBase : DINT;
    idx : DINT;
    raw : INT;
    mode : INT;
    span : REAL;
END_VAR

(* R1: 处理的通道数由 count 给出，从各数组各自的下界起算，按序号一一对应 *)
rawBase := LOWER_BOUND(analogValues, 1);
channelBase := LOWER_BOUND(channels, 1);

FOR i := 0 TO count - 1 DO
    idx := channelBase + i;
    (* R2: 只处理 enable 为 TRUE 的通道，禁用通道保持原值 *)
    IF channels[idx].enable THEN
        mode := channels[idx].measuringMode;
        raw := analogValues[rawBase + i];
        IF mode < 0 OR mode > 2 THEN
            (* R6: 非法测量模式 -> 16#8001 并跳过 *)
            channels[idx].retVal := 16#8001;
        ELSE
            IF channels[idx].hiLIM <= channels[idx].loLIM THEN
                (* R7: 量程非法 -> 16#8002 并跳过 *)
                channels[idx].retVal := 16#8002;
            ELSE
                span := channels[idx].hiLIM - channels[idx].loLIM;
                IF mode = 0 THEN
                    (* R5: 非温度线性标定 *)
                    IF channels[idx].bipolar THEN
                        (* 双极：-27648..27648 -> loLIM..hiLIM *)
                        channels[idx].outputValue := channels[idx].loLIM
                            + (INT_TO_REAL(raw) + 27648.0) * span / 55296.0;
                    ELSE
                        (* 单极：0..27648 -> loLIM..hiLIM *)
                        channels[idx].outputValue := channels[idx].loLIM
                            + INT_TO_REAL(raw) * span / 27648.0;
                    END_IF
                ELSE
                    IF mode = 1 THEN
                        (* R5: 标准温度 = raw / 10 *)
                        channels[idx].outputValue := INT_TO_REAL(raw) / 10.0;
                    ELSE
                        (* R5: 气候温度 = raw / 100 *)
                        channels[idx].outputValue := INT_TO_REAL(raw) / 100.0;
                    END_IF
                END_IF
                channels[idx].retVal := 16#0000;
            END_IF
        END_IF
    END_IF
END_FOR

(* R1: analogValues 是只读输入量，全程不被改写 *)
END_FUNCTION_BLOCK

(* ---- public-medium-03.reference.st ---- *)
FUNCTION_BLOCK FB
VAR_INPUT
    cyclicExecution : BOOL;
    trigger : BOOL;
    value : LREAL;
    windowSize : INT;
    reset : BOOL;
END_VAR
VAR_OUTPUT
    average : LREAL;
    windowSizeReached : BOOL;
    error : BOOL;
    status : WORD;
END_VAR
VAR
    buf : ARRAY[1..100] OF LREAL;
    cnt : INT;
    head : INT;
    prevTrigger : BOOL;
    trigEdge : BOOL;
    n : INT;
    i : INT;
    idx : INT;
    sum : LREAL;
    take : BOOL;
END_VAR

(* R2: 外部触发只取上升沿；周期模式与触发模式共用同一个采样标志 *)
trigEdge := trigger AND NOT prevTrigger;
prevTrigger := trigger;

(* R3: 窗口尺寸校验，16#0000 正常 / 16#8200 窗口长度错误。
   校验不受 reset 影响：尺寸非法时报错优先，避免复位把错误状态掩盖掉 *)
IF windowSize < 1 OR windowSize > 100 THEN
    error := TRUE;
    status := 16#8200;
ELSE
    error := FALSE;
    status := 16#0000;
END_IF

(* R3: 复位清空窗口统计；复位当拍不再采样，避免"清零后立刻又加一个值" *)
IF reset THEN
    cnt := 0;
    average := 0.0;
    windowSizeReached := FALSE;
ELSE
    IF NOT error THEN
        (* R1: 周期模式每扫描周期采样一次，且此模式下 trigger 无效 *)
        take := cyclicExecution OR trigEdge;
        IF take THEN
            head := head + 1;
            IF head > 100 THEN
                head := 1;
            END_IF
            buf[head] := value;
            IF cnt < 100 THEN
                cnt := cnt + 1;
            END_IF
        END_IF

        (* 窗口长度运行时可变：只对最近 n 个样本求均值，FIFO 淘汰最旧样本 *)
        n := cnt;
        IF n > windowSize THEN
            n := windowSize;
        END_IF
        windowSizeReached := cnt >= windowSize;
        IF n > 0 THEN
            sum := 0.0;
            FOR i := 0 TO n - 1 DO
                idx := head - i;
                IF idx < 1 THEN
                    idx := idx + 100;
                END_IF
                sum := sum + buf[idx];
            END_FOR
            average := sum / n;
        END_IF
    END_IF
END_IF
END_FUNCTION_BLOCK

(* ---- public-medium-04.reference.st ---- *)
FUNCTION_BLOCK FB
VAR_INPUT
    TemperatureSensorInput : REAL;
    SetTemperature : REAL;
END_VAR
VAR_OUTPUT
    CurrentTemperature : REAL;
    SetTempDisplay : REAL;
    HeaterStatus : BOOL;
    OverheatProtection : BOOL;
    HeaterOutput : BOOL;
END_VAR
VAR
    continuousHeat : TON;
    cooling : TON;
    demand : BOOL;
END_VAR

CurrentTemperature := TemperatureSensorInput;
SetTempDisplay := SetTemperature;
demand := (TemperatureSensorInput >= 0.0) AND (TemperatureSensorInput <= 100.0)
          AND (TemperatureSensorInput < SetTemperature);

cooling(IN := OverheatProtection, PT := T#3s);
IF cooling.Q THEN
    OverheatProtection := FALSE;
    cooling(IN := FALSE, PT := T#3s);
END_IF;

(* Millisecond task clock: the first representable duration over five seconds is 5001 ms. *)
continuousHeat(IN := demand AND NOT OverheatProtection, PT := T#5001ms);
IF continuousHeat.Q THEN
    OverheatProtection := TRUE;
    continuousHeat(IN := FALSE, PT := T#5001ms);
    cooling(IN := TRUE, PT := T#3s);
END_IF;
HeaterOutput := demand AND NOT OverheatProtection;
HeaterStatus := HeaterOutput;
END_FUNCTION_BLOCK

(* ---- public-medium-05.reference.st ---- *)
FUNCTION_BLOCK FB
VAR_INPUT
    Mode : BOOL;
    ForwardButton : BOOL;
    ReverseButton : BOOL;
    SensorA : BOOL;
    SensorB : BOOL;
    SensorC : BOOL;
    ButtonA : BOOL;
    ButtonB : BOOL;
    ButtonC : BOOL;
END_VAR
VAR_OUTPUT
    MotorForward : BOOL;
    MotorReverse : BOOL;
    CompletionLight : BOOL;
END_VAR
VAR
    step : INT;
END_VAR

(* R2: 正反转互锁，先无条件清零，任何分支都不允许两个方向同时输出 *)
MotorForward := FALSE;
MotorReverse := FALSE;
CompletionLight := FALSE;

IF Mode THEN
    (* R3: 自动模式按 A -> B -> C 顺序推进；
       0=等待 A，1=去 B，2=等待 B，3=去 C，4=等待 C，5=已完成 *)
    CASE step OF
        0:
            (* 必须"产品在 A（SensorA）且工位 A 加工完成（ButtonA）"才起步 *)
            IF SensorA AND ButtonA THEN
                step := 1;
                MotorForward := TRUE;
            END_IF
        1:
            (* 去 B 途中正转；B 工位传感器一到就立即停，进入等待 B *)
            MotorForward := TRUE;
            IF SensorB THEN
                MotorForward := FALSE;
                step := 2;
            END_IF
        2:
            IF SensorB AND ButtonB THEN
                step := 3;
                MotorForward := TRUE;
            END_IF
        3:
            MotorForward := TRUE;
            IF SensorC THEN
                MotorForward := FALSE;
                step := 4;
            END_IF
        4:
            (* 产品到 C 且工位 C 加工完成 -> 完成灯亮 *)
            IF SensorC AND ButtonC THEN
                CompletionLight := TRUE;
                step := 5;
            END_IF
        5:
            (* 产品被取走（SensorC 不再检测）即灭灯并回到初始等待下一件 *)
            CompletionLight := SensorC;
            IF NOT SensorC THEN
                step := 0;
            END_IF
    ELSE
        step := 0;
    END_CASE
ELSE
    (* R2: 手动模式，自动流程作废；正反转按钮互锁，两个同时按下则都不动作 *)
    step := 0;
    IF ForwardButton AND NOT ReverseButton THEN
        MotorForward := TRUE;
    END_IF
    IF ReverseButton AND NOT ForwardButton THEN
        MotorReverse := TRUE;
    END_IF
END_IF
END_FUNCTION_BLOCK

(* ---- public-medium-06.reference.st ---- *)
FUNCTION_BLOCK FB_SlabThicknessMonitor
VAR_INPUT
    THICKNESS_FAULT : BOOL;
    THICKNESS_SIGNAL_VALID : BOOL;
    CUTTING_RUN : BOOL;
    FaultTimestamp : DINT;
    CycleTime : TIME;
END_VAR
VAR_OUTPUT
    THICKNESS_ALARM : BOOL;
    Slab_Fault_Counter : UINT;
    Slab_Runtime_Accumulator : LTIME;
    Slab_Fault_History : ARRAY[0..4] OF DINT;
END_VAR
VAR
    previousFault : BOOL;
    fault : BOOL;
    remaining : TIME;
    i : INT;
END_VAR
fault := THICKNESS_SIGNAL_VALID AND THICKNESS_FAULT;
IF NOT THICKNESS_SIGNAL_VALID THEN
    remaining := T#0ms;
ELSIF fault AND NOT previousFault THEN
    remaining := T#500ms;
    IF Slab_Fault_Counter < 65535 THEN
        Slab_Fault_Counter := Slab_Fault_Counter + 1;
    END_IF;
    FOR i := 4 TO 1 BY -1 DO
        Slab_Fault_History[i] := Slab_Fault_History[i - 1];
    END_FOR;
    Slab_Fault_History[0] := FaultTimestamp;
ELSIF remaining > CycleTime THEN
    remaining := remaining - CycleTime;
ELSE
    remaining := T#0ms;
END_IF;
THICKNESS_ALARM := THICKNESS_SIGNAL_VALID AND (fault OR remaining > T#0ms);
IF CUTTING_RUN AND THICKNESS_SIGNAL_VALID AND NOT THICKNESS_FAULT THEN
    Slab_Runtime_Accumulator := Slab_Runtime_Accumulator + TIME_TO_LTIME(CycleTime);
END_IF;
previousFault := fault;
END_FUNCTION_BLOCK

(* ---- public-medium-07.reference.st ---- *)
FUNCTION_BLOCK FB_HVAC_ModeControl
VAR_INPUT
  OCCUPANCY_DETECTED : BOOL;   (* 占用检测结果（由 CO2 传感器导出） *)
  ENERGY_SAVING_MODE : BOOL;   (* TRUE=节能，FALSE=标准；只影响 Auto 模式 *)
  HVAC_MODE_SELECTOR : INT;    (* 0 Auto / 1 Comfort / 2 Economy / 3 Night *)
END_VAR
VAR_OUTPUT
  SUPPLY_FAN_RUN : BOOL;       (* 送风机运行许可 *)
  TEMP_SETPOINT_ADJUST : INT;  (* 温度设定值修正（摄氏度） *)
END_VAR
VAR
  modeValid : BOOL;            (* R1: 型号是否在合法集合 {0,1,2,3} 内 *)
  nightMode : BOOL;
  startDelay : TON;
  fanPermit : BOOL;
END_VAR

(* R1: 合法型号只有 0/1/2/3；调用方应给合法值，非法值按安全侧处理 *)
modeValid := (HVAC_MODE_SELECTOR >= 0) AND (HVAC_MODE_SELECTOR <= 3);
nightMode := HVAC_MODE_SELECTOR = 3;

fanPermit := modeValid AND OCCUPANCY_DETECTED AND NOT nightMode;
startDelay(IN := fanPermit, PT := T#30s);
SUPPLY_FAN_RUN := startDelay.Q;

(* R3 / R4 / R5 / R6: 温度设定值修正表
   - Night(3) 恒 +4，与占用无关；
   - 占用时一律 0（Night 已在上一支处理）；
   - Auto(0) 未占用：节能 +3 / 标准 +2（ENERGY_SAVING_MODE 只在这里生效）；
   - Comfort(1) 未占用 +1；Economy(2) 未占用 +4；
   - 非法型号（R1 之外）：需求未定义，按安全侧给 0。 *)
IF NOT modeValid THEN
  TEMP_SETPOINT_ADJUST := 0;
ELSIF nightMode THEN
  TEMP_SETPOINT_ADJUST := 4;
ELSIF OCCUPANCY_DETECTED THEN
  TEMP_SETPOINT_ADJUST := 0;
ELSIF HVAC_MODE_SELECTOR = 0 THEN
  IF ENERGY_SAVING_MODE THEN
    TEMP_SETPOINT_ADJUST := 3;
  ELSE
    TEMP_SETPOINT_ADJUST := 2;
  END_IF;
ELSIF HVAC_MODE_SELECTOR = 1 THEN
  TEMP_SETPOINT_ADJUST := 1;
ELSE
  TEMP_SETPOINT_ADJUST := 4;   (* Economy 未占用 *)
END_IF;

(* R6: ±4 °C 限幅；上电初值 FALSE/0 由平台默认初值保证 *)
TEMP_SETPOINT_ADJUST := LIMIT(-4, TEMP_SETPOINT_ADJUST, 4);

END_FUNCTION_BLOCK

(* ---- public-medium-08.reference.st ---- *)
(* =====================================================================
   public-medium-08  IPv4 Parsing with Format and Range Checks
   ---------------------------------------------------------------------
   平台边界（《公共题制作约定》§7）：LEN / 字符串下标 / STRING_TO_INT 可用，
   因此本解按字符扫描实现，不依赖任何 TIME 或结构体能力。

   实现约定（需求原文未逐字规定、此处显式声明的解释）：
   * 段内前导 0（"01"、"00"）按畸形处理 —— 点分十进制的规范写法里
     多位数不允许前导 0；单独一个 "0" 合法。
   * 合法点分十进制最长 15 字符（"255.255.255.255"），超长直接判非法。
   * 任何判非法的情况都把 ipValue 写成 0（需求 3）。
   ===================================================================== *)
FUNCTION_BLOCK FB_Ipv4Parser
VAR_INPUT
  ipText : STRING(254);   (* 待解析的点分十进制文本 *)
END_VAR
VAR_OUTPUT
  ipValue : UDINT;        (* 网络字节序的 32 位地址；非法输入为 0 *)
END_VAR
VAR
  s : STRING(256);        (* ipText 末尾补一个 '.'，让"最后一段"和其余段共用同一收尾逻辑 *)
  n : INT;
  i : INT;
  ch : STRING(1);
  isDigit : BOOL;
  digit : INT;
  segLen : INT;           (* 当前段已读入的数字字符数 *)
  segVal : INT;           (* 当前段的十进制值 *)
  segZeroOnly : BOOL;     (* 当前段是否"只由前导 0 开头" *)
  segCount : INT;         (* 已经收尾的段数 *)
  segments : ARRAY[0..3] OF INT;
  ok : BOOL;              (* 合法性结论（内部观察量） *)
  run : BOOL;
END_VAR

s := CONCAT(ipText, '.');
n := LEN(s);
ok := TRUE;
segCount := 0;
segLen := 0;
segVal := 0;
segZeroOnly := FALSE;

(* R1 / R3: 合法点分十进制最长 15 字符；超长直接判非法 *)
IF LEN(ipText) > 15 THEN
  ok := FALSE;
END_IF;

(* R1: 逐字符扫描，'.' 收尾一段，其余必须是十进制数字 *)
FOR i := 1 TO 16 DO
  run := ok AND (i <= n);
  IF run THEN
    ch := s[i];
    isDigit := (ch >= '0') AND (ch <= '9');
    IF ch = '.' THEN
      IF segLen = 0 THEN
        ok := FALSE;            (* R3: 空段（空输入 / 连续点 / 以点结尾） *)
      ELSIF segLen > 3 THEN
        ok := FALSE;            (* R3: 段内数字超过 3 位 *)
      ELSIF segVal > 255 THEN
        ok := FALSE;            (* R3: 段值超出 0~255 *)
      ELSIF segCount > 3 THEN
        ok := FALSE;            (* R3: 段数超过 4 *)
      ELSE
        segments[segCount] := segVal;
        segCount := segCount + 1;
      END_IF;
      segLen := 0;
      segVal := 0;
      segZeroOnly := FALSE;
    ELSIF isDigit THEN
      digit := STRING_TO_INT(ch);
      IF (segLen = 0) AND (digit = 0) THEN
        segZeroOnly := TRUE;    (* 段首是 0：只允许单独一个 "0" *)
      ELSIF segZeroOnly THEN
        ok := FALSE;            (* R3: 前导 0（"01"/"00"）视为畸形 *)
      END_IF;
      IF segLen < 3 THEN
        segLen := segLen + 1;
        segVal := segVal * 10 + digit;
      ELSE
        segLen := 4;            (* 超过 3 位，留到收尾分支判非法 *)
      END_IF;
    ELSE
      ok := FALSE;              (* R3: 非数字、非点字符（空格、字母、符号…） *)
    END_IF;
  END_IF;
END_FOR;

(* R1 / R3: 必须恰好四段 *)
IF ok AND (segCount <> 4) THEN
  ok := FALSE;
END_IF;

(* R2: 网络字节序拼装（第一段占最高 8 位）；R3: 非法输入 → 0（0.0.0.0 也是 0） *)
ipValue := 0;
IF ok THEN
  FOR i := 0 TO 3 DO
    ipValue := ipValue * 256 + segments[i];
  END_FOR;
END_IF;

END_FUNCTION_BLOCK
